(* CODESYS project NavBar.xml

Project tree, tasks and I/O mapping:
  visualisation NavBar
*)

// /NavBar
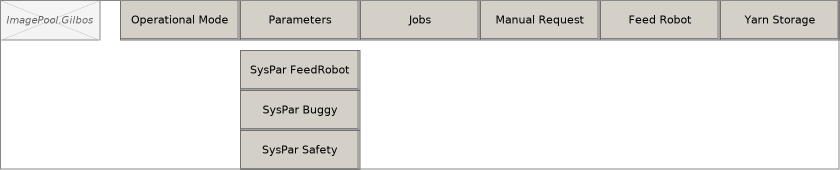
VISUALIZATION NavBar  // 840x170
    Button (120,0 120x40), "Operational Mode"
        tap GVL_Project.fbProject._fbNavBarController._btnOperationalMode.xbtn
    Image (0,0 100x40), image: ImagePool.Gilbos
    Button (240,0 120x40), "Parameters"
        tap GVL_Project.fbProject._fbNavBarController._btnParameters.xbtn p1329445385=TRUE
        OnMouseEnter: execute { GVL_Project.fbProject._fbNavBarController.xHoverParameters := TRUE; }
        OnMouseLeave: execute { GVL_Project.fbProject._fbNavBarController.xHoverParameters := FALSE; }
    Button (360,0 120x40), "Jobs"
        tap GVL_Project.fbProject._fbNavBarController._btnJobManager.xbtn
    Button (240,50 120x40), "SysPar FeedRobot", invisible if: GVL_Project.fbProject._fbNavBarController.xHideParameters
        tap GVL_Project.fbProject._fbNavBarController._btnSysParFR.xbtn
        OnMouseEnter: execute { GVL_Project.fbProject._fbNavBarController.xHoverParameters := TRUE; }
        OnMouseLeave: execute { GVL_Project.fbProject._fbNavBarController.xHoverParameters := FALSE; }
    Button (240,90 120x40), "SysPar Buggy", invisible if: GVL_Project.fbProject._fbNavBarController.xHideParameters
        tap GVL_Project.fbProject._fbNavBarController._btnSysParBuggy.xbtn
        OnMouseEnter: execute { GVL_Project.fbProject._fbNavBarController.xHoverParameters := TRUE; }
        OnMouseLeave: execute { GVL_Project.fbProject._fbNavBarController.xHoverParameters := FALSE; }
    Button (480,0 120x40), "Manual Request"
        tap GVL_Project.fbProject._fbNavBarController._btnManualRequest.xbtn
    Button (600,0 120x40), "Feed Robot"
        tap GVL_Project.fbProject._fbNavBarController._btnFeedRobot.xbtn
    Button (720,0 120x40), "Yarn Storage"
        tap GVL_Project.fbProject._fbNavBarController._btnYarnStorage.xbtn
    Button (240,130 120x40), "SysPar Safety", invisible if: GVL_Project.fbProject._fbNavBarController.xHideParameters
        tap GVL_Project.fbProject._fbNavBarController._btnSysParSafety.xbtn
        OnMouseEnter: execute { GVL_Project.fbProject._fbNavBarController.xHoverParameters := TRUE; }
        OnMouseLeave: execute { GVL_Project.fbProject._fbNavBarController.xHoverParameters := FALSE; }
END_VISUALIZATION
